Fanuc KAREL source: KB00017.KL

PROGRAM KB00017
%NOLOCKGROUP
%ENVIRONMENT UIF
VAR
  P1: STRING[80]
  P2: STRING[80]
  P3: INTEGER
BEGIN
  P1 = 'A'
  P2 = 'A'
  P3 = 1
  CHECK_DICT(P1, P2, P3)
END KB00017
